FUNCTION_BLOCK FB_ZylinderAuslauf
VAR_INPUT
END_VAR
VAR_OUTPUT
END_VAR
VAR
END_VAR

GVL_IO.xVentilAuslaufAS := GVL_IO.xWeicheAcceptBereit;
GVL_IO.xVentilAuslaufGS := NOT GVL_IO.xWeicheAcceptBereit;

GVL_IO.xZylinderAuslaufBereit := GVL_IO.xZylinderAuslaufAS;

END_FUNCTION_BLOCK

(* stored: Version 1.1.0.1
   POU FB_ZylinderAuslauf: Id {89dcefb7-7762-4274-8ce3-5883557cf7f7}, SpecialFunc None *)
